(* PLC project Mixer, Beremiz Mixer 1 *)
(* stored: creationDateTime 2026-10-19T10:00:00, modificationDateTime 2026-10-19T10:00:00 *)

TYPE E_Mode : (Idle, Fill := 10, Mix);
END_TYPE

TYPE ST_Tank : STRUCT
  Level : REAL;
  Name : STRING(20) := 'Tank A';
  History : ARRAY[0..9] OF INT;
END_STRUCT;
END_TYPE

TYPE T_Percent : INT(0..100);
END_TYPE

FUNCTION Scale : REAL
  VAR_INPUT
    Raw : INT;
  END_VAR

Scale := INT_TO_REAL(Raw) / 27.648;
END_FUNCTION

FUNCTION_BLOCK Counter
  VAR_INPUT
    Reset : BOOL;
  END_VAR
  VAR_OUTPUT
    OUT : INT;
  END_VAR
  VAR
    Cnt : INT;
  END_VAR

(* FBD diagram, written out as Structured Text *)
Cnt := SEL(Reset, 1 + Cnt, 0);
OUT := Cnt;
END_FUNCTION_BLOCK

PROGRAM Main
  VAR_INPUT
    Start : BOOL;
    Stop : BOOL;
    Level : INT;
  END_VAR
  VAR_OUTPUT
    Motor : BOOL;
    Alarm : BOOL;
  END_VAR
  VAR
    Delay : TON;
    Cycles : Counter;
    Mode : E_Mode := E_Mode.Idle;
  END_VAR
  VAR  (* added by the conversion: wires and edge detectors of the diagram *)
    R_TRIG1 : R_TRIG;
  END_VAR

(* LD diagram, written out as Structured Text *)
Motor := (Start OR Motor) AND NOT Stop;
R_TRIG1(CLK := Motor);
Delay(IN := R_TRIG1.Q, PT := T#5s);
IF Delay.Q THEN Alarm := TRUE; END_IF;
END_PROGRAM

PROGRAM Sequence
  VAR_INPUT
    Go : BOOL;
    Done : BOOL;
  END_VAR
  VAR_OUTPUT
    Valve : BOOL;
    Pump : BOOL;
  END_VAR

INITIAL_STEP Init:
END_STEP
TRANSITION FROM Init TO Filling
  := Go AND NOT Done;
END_TRANSITION
STEP Filling:
  OpenValve(N);
  FILLING_INLINE1(S);
END_STEP
ACTION FILLING_INLINE1:
  Pump := TRUE;
END_ACTION
TRANSITION FROM Filling TO Init  (* Finished *)
  := Done;
END_TRANSITION
TRANSITION FROM Filling TO Init
  := NOT Go;
END_TRANSITION

ACTION OpenValve:
Valve := TRUE;
END_ACTION
END_PROGRAM

CONFIGURATION config
  RESOURCE cpu ON PLC
    VAR_GLOBAL
      Setpoint : REAL := 42.5;
    END_VAR
    TASK fast(INTERVAL := T#10ms, PRIORITY := 1);
    TASK slow(INTERVAL := T#100ms, PRIORITY := 5);
    PROGRAM main_inst WITH fast : Main;
    PROGRAM seq_inst WITH slow : Sequence;
  END_RESOURCE
END_CONFIGURATION
